(* IEC 61131-3 sources: BODAS-HelloWorld/st/bodas_rc18_12_40/plc_logic/application/03_privatelibrary/datatypes/maintask, 6 files *)

(* ---- enu_listctrlvlv-enu_listCtrlVlv.st ---- *)
(* --- Interface --- *)
{attribute 'qualified_only'}
{attribute 'strict'}
TYPE enu_ListCtrlVlv : (
		st_fctOff_cenu := 0, (* Default value *)
		st_fctOnPos_cenu,
		st_fctOnNeg_cenu
	);
END_TYPE

(* ---- enu_maintaskstate-enu_MainTaskState.st ---- *)
(* --- Interface --- *)
{attribute 'qualified_only'}
{attribute 'strict'}
TYPE enu_MainTaskState :
(
	MT_INIT := 0,
	MT_CYCLE
);
END_TYPE

(* ---- struc_dbgmgrprm-struc_DbgMgrPrm.st ---- *)
(* --- Interface --- *)
TYPE struc_DbgMgrPrm : STRUCT
		flgXcpOn_b          : BOOL;
		flgStoreDataToNvm_b : BOOL;
	END_STRUCT
END_TYPE

(* ---- struc_errmemmgr_prevactvdfes-struc_ErrMemMgr_prevActvDfes.st ---- *)
(* --- Interface --- *)
TYPE struc_ErrMemMgr_prevActvDfes : STRUCT
		idxPrevActvDfes_u32 : UDINT; (* DTC OF previously active/deactive error in DFES *)
		tiStamp_min_u32     : UDINT; (* TIME stamp when DFES got previously active *)
	END_STRUCT
END_TYPE

(* ---- struc_mnginhb-struc_MngInhb.st ---- *)
(* --- Interface --- *)
TYPE struc_MngInhb : STRUCT
		st_flgUBattLowDetd_b : BOOL;
		st_flgInhbActv_b     : BOOL;
		st_flgOutpLockd_b    : BOOL;
		UBatt_mV_u16         : UINT;
		NrCycDebRst_u16      : UINT;
	END_STRUCT
END_TYPE

(* ---- struc_para-struc_para.st ---- *)
(* --- Interface --- *)
TYPE struc_para : STRUCT
		fctPmp_s16       : INT;
		listCtrlVlv_enu  : enu_listCtrlVlv; (* parameter DID 0xC002, list {0 - Off; 1 - OnPos; 2 - OnNeg;} *)
		nrCogs_s16       : INT;
		iSpSafout1_u16   : UINT;
		iSpSafout2_u16   : UINT;
		nEngSpd_rpm_au16 : ARRAY[0..2] OF UINT;
		eff_perc_au16    : ARRAY[0..2] OF UINT;
		PrmDbg_struc     : struc_DbgMgrPrm;
	END_STRUCT
END_TYPE
